TYPE "ST_TwoHandHal"
VERSION : 0.1
   STRUCT
      LeftPressed : Bool;
      RightPressed : Bool;
      SafeActive : Bool;
      FieldbusHealthy : Bool;
   END_STRUCT;

END_TYPE

